Staubli VAL3: HMI_FrameSet.dtx

mdesc mNomSpeed = {accel=25, vel=50, decel=25, leave=0, reach=0, blend=off}
string sFrameList
string sToolList
string sSelFrame
string sSelTool
bool bBool[6]
bool bBack
public num nTool[6]
bool bModifyTool
bool bCancelTool
num nFrame[6]
bool bModifyFrame
bool bCancelFrame
string sUsingTool
string sUsingFrame
num nNmbValue[6]
num nWizardStep
bool bPrevious
bool bTeach
bool bMove
bool bNext
string sLastTool
tool tUsingTool = {fatherId=flange[0]}
string sTitle
num _nTool
